(* IEC 61131-3 sources: sis-interlock-demo/pytests/golden/mini/tests/POUs/Generated/FB_CemGen01_Test, 24 files *)

(* ---- FB_CemGen01_Test.decl.st ---- *)
// AUTO-GENERATED by cemgen 1.0.0 — не редактировать: правьте матрицу и запустите
//   python -m cemgen generate <файл матрицы .csv или .xlsx>
// Матрица: TEST-U301-CEM, объект U-301, ревизия 1 от 2026-10-16, SHA-256 сетки 9067fda96ae55e67
// Назначение: набор coUnit: сценарии по матрице TEST-U301-CEM, тесты 1–24 (DESIGN.md, 12.4).
//             Ожидаемые значения — эталонная модель cemgen. Стенд FB_SisHarness — по экземпляру на
//             тест.
// Автор:      pytest; код — генератор cemgen
// Версия:     1.0.0
// Документ:   docs/DESIGN.md, раздел «10. Генератор cemgen»; docs/cause_effect_matrix.md
// ВНИМАНИЕ:   код демонстрационный и не предназначен для систем безопасности. Реальная ПАЗ требует
//             определения SIL, сертифицированных аппаратных и программных средств и валидации по
//             ГОСТ Р МЭК 61511.
FUNCTION_BLOCK FB_CemGen01_Test EXTENDS coUnit.FB_TestSuite
VAR
    fbH001 : FB_SisHarness;   // Matrix_TSH301Demand_TripsOwnEffects
    fbH002 : FB_SisHarness;   // Matrix_TSH301Delay_TripsExactlyAtDelay
    fbH003 : FB_SisHarness;   // Matrix_TSH301Override_Denied
    fbH004 : FB_SisHarness;   // Matrix_TSH301Reset_OnlyAfterClear
    fbH005 : FB_SisHarness;   // Matrix_TSH301ChannelInvalid_MatchesPolicy
    fbH006 : FB_SisHarness;   // Matrix_TSH301Bypass_Denied
    fbH007 : FB_SisHarness;   // Matrix_PSL302Demand_TripsOwnEffects
    fbH008 : FB_SisHarness;   // Matrix_PSL302Override_ExpiresThenTrips
    fbH009 : FB_SisHarness;   // Matrix_PSL302Override_ClearsAfterConfirm
    fbH010 : FB_SisHarness;   // Matrix_PSL302Override_DemandBackRestartsConfirm
    fbH011 : FB_SisHarness;   // Matrix_PSL302Override_ExpiryBoundsConfirm
    fbH012 : FB_SisHarness;   // Matrix_PSL302Reset_OnlyAfterClear
    fbH013 : FB_SisHarness;   // Matrix_PSL302ChannelInvalid_MatchesPolicy
    fbH014 : FB_SisHarness;   // Matrix_PSL302Bypass_ExpiresBackToVoting
    fbH015 : FB_SisHarness;   // Matrix_XS303Demand_TripsOwnEffects
    fbH016 : FB_SisHarness;   // Matrix_XS303Delay_TripsExactlyAtDelay
    fbH017 : FB_SisHarness;   // Matrix_XS303Override_Denied
    fbH018 : FB_SisHarness;   // Matrix_XS303Reset_OnlyAfterClear
    fbH019 : FB_SisHarness;   // Matrix_FirstOutTSH301ThenPSL302_RecordsFirst
    fbH020 : FB_SisHarness;   // Matrix_FirstOutPSL302ThenXS303_RecordsFirst
    fbH021 : FB_SisHarness;   // Matrix_FirstOutXS303ThenTSH301_RecordsFirst
    fbH022 : FB_SisHarness;   // Matrix_Start_EnergizedWithoutReset
    fbH023 : FB_SisHarness;   // Matrix_FirstOutSimultaneous_LowestIndex
    fbH024 : FB_SisHarness;   // Matrix_GeneratedCfg_PassesChecks
END_VAR

(* ---- FirstOutPSL302ThenXS303RecordsFirst.method.decl.st ---- *)
// AUTO-GENERATED by cemgen 1.0.0 — не редактировать: правьте матрицу и запустите
//   python -m cemgen generate <файл матрицы .csv или .xlsx>
// Матрица: TEST-U301-CEM, объект U-301, ревизия 1 от 2026-10-16, SHA-256 сетки 9067fda96ae55e67
// Назначение: тест Matrix_FirstOutPSL302ThenXS303_RecordsFirst набора FB_CemGen01_Test (сценарий по
//             матрице, DESIGN.md, 12.4).
// Автор:      pytest; код — генератор cemgen
// Версия:     1.0.0
// Документ:   docs/DESIGN.md, раздел «10. Генератор cemgen»; docs/cause_effect_matrix.md
// ВНИМАНИЕ:   код демонстрационный и не предназначен для систем безопасности. Реальная ПАЗ требует
//             определения SIL, сертифицированных аппаратных и программных средств и валидации по
//             ГОСТ Р МЭК 61511.
// Первопричина: требование PSL302, фиксация через 0 с; затем требование XS303, фиксация через 500 мс →
// первопричина PSL302, в маске первопричины только PSL302, ltFirstOut — момент фиксации PSL302, XS303
// — среди зафиксированных.
METHOD PRIVATE FirstOutPSL302ThenXS303RecordsFirst
VAR
    xArmed : BOOL;    // стенд взведён: все следствия под напряжением после сброса
    ltT0   : LTIME;   // момент t0 по подменному времени стенда
END_VAR

(* ---- FirstOutSimultaneousLowestIndex.method.decl.st ---- *)
// AUTO-GENERATED by cemgen 1.0.0 — не редактировать: правьте матрицу и запустите
//   python -m cemgen generate <файл матрицы .csv или .xlsx>
// Матрица: TEST-U301-CEM, объект U-301, ревизия 1 от 2026-10-16, SHA-256 сетки 9067fda96ae55e67
// Назначение: тест Matrix_FirstOutSimultaneous_LowestIndex набора FB_CemGen01_Test (сценарий по
//             матрице, DESIGN.md, 12.4).
// Автор:      pytest; код — генератор cemgen
// Версия:     1.0.0
// Документ:   docs/DESIGN.md, раздел «10. Генератор cemgen»; docs/cause_effect_matrix.md
// ВНИМАНИЕ:   код демонстрационный и не предназначен для систем безопасности. Реальная ПАЗ требует
//             определения SIL, сертифицированных аппаратных и программных средств и валидации по
//             ГОСТ Р МЭК 61511.
// Одновременная фиксация TSH301 и PSL302 (без общих каналов) в одном вызове: требования подаются со
// сдвигом на разницу задержек → первопричина — младшая причина, в маске первопричины обе.
METHOD PRIVATE FirstOutSimultaneousLowestIndex
VAR
    xArmed : BOOL;   // стенд взведён: все следствия под напряжением после сброса
END_VAR

(* ---- FirstOutTSH301ThenPSL302RecordsFirst.method.decl.st ---- *)
// AUTO-GENERATED by cemgen 1.0.0 — не редактировать: правьте матрицу и запустите
//   python -m cemgen generate <файл матрицы .csv или .xlsx>
// Матрица: TEST-U301-CEM, объект U-301, ревизия 1 от 2026-10-16, SHA-256 сетки 9067fda96ae55e67
// Назначение: тест Matrix_FirstOutTSH301ThenPSL302_RecordsFirst набора FB_CemGen01_Test (сценарий
//             по матрице, DESIGN.md, 12.4).
// Автор:      pytest; код — генератор cemgen
// Версия:     1.0.0
// Документ:   docs/DESIGN.md, раздел «10. Генератор cemgen»; docs/cause_effect_matrix.md
// ВНИМАНИЕ:   код демонстрационный и не предназначен для систем безопасности. Реальная ПАЗ требует
//             определения SIL, сертифицированных аппаратных и программных средств и валидации по
//             ГОСТ Р МЭК 61511.
// Первопричина: требование TSH301, фиксация через 1 с; затем требование PSL302, фиксация через 0 с →
// первопричина TSH301, в маске первопричины только TSH301, ltFirstOut — момент фиксации TSH301, PSL302
// — среди зафиксированных.
METHOD PRIVATE FirstOutTSH301ThenPSL302RecordsFirst
VAR
    xArmed : BOOL;    // стенд взведён: все следствия под напряжением после сброса
    ltT0   : LTIME;   // момент t0 по подменному времени стенда
END_VAR

(* ---- FirstOutXS303ThenTSH301RecordsFirst.method.decl.st ---- *)
// AUTO-GENERATED by cemgen 1.0.0 — не редактировать: правьте матрицу и запустите
//   python -m cemgen generate <файл матрицы .csv или .xlsx>
// Матрица: TEST-U301-CEM, объект U-301, ревизия 1 от 2026-10-16, SHA-256 сетки 9067fda96ae55e67
// Назначение: тест Matrix_FirstOutXS303ThenTSH301_RecordsFirst набора FB_CemGen01_Test (сценарий по
//             матрице, DESIGN.md, 12.4).
// Автор:      pytest; код — генератор cemgen
// Версия:     1.0.0
// Документ:   docs/DESIGN.md, раздел «10. Генератор cemgen»; docs/cause_effect_matrix.md
// ВНИМАНИЕ:   код демонстрационный и не предназначен для систем безопасности. Реальная ПАЗ требует
//             определения SIL, сертифицированных аппаратных и программных средств и валидации по
//             ГОСТ Р МЭК 61511.
// Первопричина: требование XS303, фиксация через 500 мс; затем требование TSH301, фиксация через 1 с →
// первопричина XS303, в маске первопричины только XS303, ltFirstOut — момент фиксации XS303, TSH301 —
// среди зафиксированных.
METHOD PRIVATE FirstOutXS303ThenTSH301RecordsFirst
VAR
    xArmed : BOOL;    // стенд взведён: все следствия под напряжением после сброса
    ltT0   : LTIME;   // момент t0 по подменному времени стенда
END_VAR

(* ---- GeneratedCfgPassesChecks.method.decl.st ---- *)
// AUTO-GENERATED by cemgen 1.0.0 — не редактировать: правьте матрицу и запустите
//   python -m cemgen generate <файл матрицы .csv или .xlsx>
// Матрица: TEST-U301-CEM, объект U-301, ревизия 1 от 2026-10-16, SHA-256 сетки 9067fda96ae55e67
// Назначение: тест Matrix_GeneratedCfg_PassesChecks набора FB_CemGen01_Test (сценарий по матрице,
//             DESIGN.md, 12.4).
// Автор:      pytest; код — генератор cemgen
// Версия:     1.0.0
// Документ:   docs/DESIGN.md, раздел «10. Генератор cemgen»; docs/cause_effect_matrix.md
// ВНИМАНИЕ:   код демонстрационный и не предназначен для систем безопасности. Реальная ПАЗ требует
//             определения SIL, сертифицированных аппаратных и программных средств и валидации по
//             ГОСТ Р МЭК 61511.
// Сгенерированная конфигурация: F_CemCrc(CEM_CFG) = 16#0F15 = CEM_CFG.wMatrixCrc, F_CemCheckCfg без
// ошибок; после взвода нет ошибок конфигурации у матрицы и у групп голосования.
METHOD PRIVATE GeneratedCfgPassesChecks
VAR
    stCfg  : ST_CemCfg;      // копия GVL_SisCfg.CEM_CFG
    wCrc   : WORD;           // CRC сгенерированной матрицы
    wErr   : WORD;           // биты ошибок конфигурации матрицы
    xArmed : BOOL;           // стенд взведён: все следствия под напряжением после сброса
    stVs   : ST_VotingSts;   // копия состояния группы голосования
END_VAR

(* ---- PSL302BypassExpiresBackToVoting.method.decl.st ---- *)
// AUTO-GENERATED by cemgen 1.0.0 — не редактировать: правьте матрицу и запустите
//   python -m cemgen generate <файл матрицы .csv или .xlsx>
// Матрица: TEST-U301-CEM, объект U-301, ревизия 1 от 2026-10-16, SHA-256 сетки 9067fda96ae55e67
// Назначение: тест Matrix_PSL302Bypass_ExpiresBackToVoting набора FB_CemGen01_Test (сценарий по
//             матрице, DESIGN.md, 12.4).
// Автор:      pytest; код — генератор cemgen
// Версия:     1.0.0
// Документ:   docs/DESIGN.md, раздел «10. Генератор cemgen»; docs/cause_effect_matrix.md
// ВНИМАНИЕ:   код демонстрационный и не предназначен для систем безопасности. Реальная ПАЗ требует
//             определения SIL, сертифицированных аппаратных и программных средств и валидации по
//             ГОСТ Р МЭК 61511.
// Причина 2 PSL302: ключ разрешения байпасов, байпас PS302A → Active; канал недостоверен → Bypassed,
// не сработало; на t0 + 1 ч − шаг — Active; ровно на t0 + 1 ч — Expired, BypassExpired, канал Invalid;
// далее — по эталонной модели.
METHOD PRIVATE PSL302BypassExpiresBackToVoting
VAR
    xArmed : BOOL;           // стенд взведён: все следствия под напряжением после сброса
    stVs   : ST_VotingSts;   // копия состояния группы голосования
END_VAR

(* ---- PSL302ChannelInvalidMatchesPolicy.method.decl.st ---- *)
// AUTO-GENERATED by cemgen 1.0.0 — не редактировать: правьте матрицу и запустите
//   python -m cemgen generate <файл матрицы .csv или .xlsx>
// Матрица: TEST-U301-CEM, объект U-301, ревизия 1 от 2026-10-16, SHA-256 сетки 9067fda96ae55e67
// Назначение: тест Matrix_PSL302ChannelInvalid_MatchesPolicy набора FB_CemGen01_Test (сценарий по
//             матрице, DESIGN.md, 12.4).
// Автор:      pytest; код — генератор cemgen
// Версия:     1.0.0
// Документ:   docs/DESIGN.md, раздел «10. Генератор cemgen»; docs/cause_effect_matrix.md
// ВНИМАНИЕ:   код демонстрационный и не предназначен для систем безопасности. Реальная ПАЗ требует
//             определения SIL, сертифицированных аппаратных и программных средств и валидации по
//             ГОСТ Р МЭК 61511.
// Причина 2 PSL302 (2oo2, VoteTrip): канал PS302A недостоверен → действующая схема и срабатывание по
// политике деградации; если не сработало — требование на PS302B → по эталонной модели.
METHOD PRIVATE PSL302ChannelInvalidMatchesPolicy
VAR
    xArmed : BOOL;           // стенд взведён: все следствия под напряжением после сброса
    stVs   : ST_VotingSts;   // копия состояния группы голосования
END_VAR

(* ---- PSL302DemandTripsOwnEffects.method.decl.st ---- *)
// AUTO-GENERATED by cemgen 1.0.0 — не редактировать: правьте матрицу и запустите
//   python -m cemgen generate <файл матрицы .csv или .xlsx>
// Матрица: TEST-U301-CEM, объект U-301, ревизия 1 от 2026-10-16, SHA-256 сетки 9067fda96ae55e67
// Назначение: тест Matrix_PSL302Demand_TripsOwnEffects набора FB_CemGen01_Test (сценарий по
//             матрице, DESIGN.md, 12.4).
// Автор:      pytest; код — генератор cemgen
// Версия:     1.0.0
// Документ:   docs/DESIGN.md, раздел «10. Генератор cemgen»; docs/cause_effect_matrix.md
// ВНИМАНИЕ:   код демонстрационный и не предназначен для систем безопасности. Реальная ПАЗ требует
//             определения SIL, сертифицированных аппаратных и программных средств и валидации по
//             ГОСТ Р МЭК 61511.
// Причина 2 PSL302 (2oo2, задержка 0 с): требование PS302A, PS302B = 0 отключает XV301, M302;
// остальные следствия под напряжением; первопричина PSL302.
METHOD PRIVATE PSL302DemandTripsOwnEffects
VAR
    xArmed : BOOL;   // стенд взведён: все следствия под напряжением после сброса
END_VAR

(* ---- PSL302OverrideClearsAfterConfirm.method.decl.st ---- *)
// AUTO-GENERATED by cemgen 1.0.0 — не редактировать: правьте матрицу и запустите
//   python -m cemgen generate <файл матрицы .csv или .xlsx>
// Матрица: TEST-U301-CEM, объект U-301, ревизия 1 от 2026-10-16, SHA-256 сетки 9067fda96ae55e67
// Назначение: тест Matrix_PSL302Override_ClearsAfterConfirm набора FB_CemGen01_Test (сценарий по
//             матрице, DESIGN.md, 12.4).
// Автор:      pytest; код — генератор cemgen
// Версия:     1.0.0
// Документ:   docs/DESIGN.md, раздел «10. Генератор cemgen»; docs/cause_effect_matrix.md
// ВНИМАНИЕ:   код демонстрационный и не предназначен для систем безопасности. Реальная ПАЗ требует
//             определения SIL, сертифицированных аппаратных и программных средств и валидации по
//             ГОСТ Р МЭК 61511.
// Причина 2 PSL302: пусковой обход и требование в t0; норма с t1 = t0 + шаг; на t1 + 30 с − шаг обход
// действует; ровно на t1 + 30 с (подтверждение нормы) — OverrideCleared, обхода нет, причина не
// зафиксирована, следствия под напряжением (R-12).
METHOD PRIVATE PSL302OverrideClearsAfterConfirm
VAR
    xArmed : BOOL;   // стенд взведён: все следствия под напряжением после сброса
END_VAR

(* ---- PSL302OverrideDemandBackRestartsConfirm.method.decl.st ---- *)
// AUTO-GENERATED by cemgen 1.0.0 — не редактировать: правьте матрицу и запустите
//   python -m cemgen generate <файл матрицы .csv или .xlsx>
// Матрица: TEST-U301-CEM, объект U-301, ревизия 1 от 2026-10-16, SHA-256 сетки 9067fda96ae55e67
// Назначение: тест Matrix_PSL302Override_DemandBackRestartsConfirm набора FB_CemGen01_Test
//             (сценарий по матрице, DESIGN.md, 12.4).
// Автор:      pytest; код — генератор cemgen
// Версия:     1.0.0
// Документ:   docs/DESIGN.md, раздел «10. Генератор cemgen»; docs/cause_effect_matrix.md
// ВНИМАНИЕ:   код демонстрационный и не предназначен для систем безопасности. Реальная ПАЗ требует
//             определения SIL, сертифицированных аппаратных и программных средств и валидации по
//             ГОСТ Р МЭК 61511.
// Причина 2 PSL302: пусковой обход и требование в t0; норма с t1; ровно на t1 + 30 с, когда обход
// снялся бы, требование снова — обход действует, подтверждение нормы сброшено; норма с t2; на t2 + 30
// с − шаг обход действует; на t2 + 30 с — OverrideCleared.
METHOD PRIVATE PSL302OverrideDemandBackRestartsConfirm
VAR
    xArmed : BOOL;   // стенд взведён: все следствия под напряжением после сброса
END_VAR

(* ---- PSL302OverrideExpiresThenTrips.method.decl.st ---- *)
// AUTO-GENERATED by cemgen 1.0.0 — не редактировать: правьте матрицу и запустите
//   python -m cemgen generate <файл матрицы .csv или .xlsx>
// Матрица: TEST-U301-CEM, объект U-301, ревизия 1 от 2026-10-16, SHA-256 сетки 9067fda96ae55e67
// Назначение: тест Matrix_PSL302Override_ExpiresThenTrips набора FB_CemGen01_Test (сценарий по
//             матрице, DESIGN.md, 12.4).
// Автор:      pytest; код — генератор cemgen
// Версия:     1.0.0
// Документ:   docs/DESIGN.md, раздел «10. Генератор cemgen»; docs/cause_effect_matrix.md
// ВНИМАНИЕ:   код демонстрационный и не предназначен для систем безопасности. Реальная ПАЗ требует
//             определения SIL, сертифицированных аппаратных и программных средств и валидации по
//             ГОСТ Р МЭК 61511.
// Причина 2 PSL302: ключ разрешения обходов, запрос пускового обхода и требование в одном вызове t0;
// до t0 + 10 мин − шаг обход действует, причина не зафиксирована; ровно на t0 + 10 мин —
// OverrideExpired, фиксация, первопричина PSL302.
METHOD PRIVATE PSL302OverrideExpiresThenTrips
VAR
    xArmed : BOOL;   // стенд взведён: все следствия под напряжением после сброса
END_VAR

(* ---- PSL302OverrideExpiryBoundsConfirm.method.decl.st ---- *)
// AUTO-GENERATED by cemgen 1.0.0 — не редактировать: правьте матрицу и запустите
//   python -m cemgen generate <файл матрицы .csv или .xlsx>
// Матрица: TEST-U301-CEM, объект U-301, ревизия 1 от 2026-10-16, SHA-256 сетки 9067fda96ae55e67
// Назначение: тест Matrix_PSL302Override_ExpiryBoundsConfirm набора FB_CemGen01_Test (сценарий по
//             матрице, DESIGN.md, 12.4).
// Автор:      pytest; код — генератор cemgen
// Версия:     1.0.0
// Документ:   docs/DESIGN.md, раздел «10. Генератор cemgen»; docs/cause_effect_matrix.md
// ВНИМАНИЕ:   код демонстрационный и не предназначен для систем безопасности. Реальная ПАЗ требует
//             определения SIL, сертифицированных аппаратных и программных средств и валидации по
//             ГОСТ Р МЭК 61511.
// Причина 2 PSL302: пусковой обход и требование в t0; норма с t0 + 9 мин 30 с + шаг — подтверждение
// (30 с) закончилось бы после срока; на t0 + 10 мин − шаг обход действует; ровно на t0 + 10 мин —
// OverrideExpired (срок — верхняя граница), OverrideCleared нет, причина не зафиксирована (требования
// нет).
METHOD PRIVATE PSL302OverrideExpiryBoundsConfirm
VAR
    xArmed : BOOL;   // стенд взведён: все следствия под напряжением после сброса
END_VAR

(* ---- PSL302ResetOnlyAfterClear.method.decl.st ---- *)
// AUTO-GENERATED by cemgen 1.0.0 — не редактировать: правьте матрицу и запустите
//   python -m cemgen generate <файл матрицы .csv или .xlsx>
// Матрица: TEST-U301-CEM, объект U-301, ревизия 1 от 2026-10-16, SHA-256 сетки 9067fda96ae55e67
// Назначение: тест Matrix_PSL302Reset_OnlyAfterClear набора FB_CemGen01_Test (сценарий по матрице,
//             DESIGN.md, 12.4).
// Автор:      pytest; код — генератор cemgen
// Версия:     1.0.0
// Документ:   docs/DESIGN.md, раздел «10. Генератор cemgen»; docs/cause_effect_matrix.md
// ВНИМАНИЕ:   код демонстрационный и не предназначен для систем безопасности. Реальная ПАЗ требует
//             определения SIL, сертифицированных аппаратных и программных средств и валидации по
//             ГОСТ Р МЭК 61511.
// Причина 2 PSL302: срабатывание; сброс при требовании → ResetDenied, блокирует PSL302, следствия
// обесточены; норма → следствия всё ещё обесточены (фиксация); сброс → все следствия под напряжением.
METHOD PRIVATE PSL302ResetOnlyAfterClear
VAR
    xArmed : BOOL;          // стенд взведён: все следствия под напряжением после сброса
    stEv   : ST_SisEvent;   // последнее событие журнала
END_VAR

(* ---- TSH301BypassDenied.method.decl.st ---- *)
// AUTO-GENERATED by cemgen 1.0.0 — не редактировать: правьте матрицу и запустите
//   python -m cemgen generate <файл матрицы .csv или .xlsx>
// Матрица: TEST-U301-CEM, объект U-301, ревизия 1 от 2026-10-16, SHA-256 сетки 9067fda96ae55e67
// Назначение: тест Matrix_TSH301Bypass_Denied набора FB_CemGen01_Test (сценарий по матрице,
//             DESIGN.md, 12.4).
// Автор:      pytest; код — генератор cemgen
// Версия:     1.0.0
// Документ:   docs/DESIGN.md, раздел «10. Генератор cemgen»; docs/cause_effect_matrix.md
// ВНИМАНИЕ:   код демонстрационный и не предназначен для систем безопасности. Реальная ПАЗ требует
//             определения SIL, сертифицированных аппаратных и программных средств и валидации по
//             ГОСТ Р МЭК 61511.
// Причина 1 TSH301: байпас запрещён (bypass_max = 0); ключ разрешения байпасов, запрос байпаса TT301 →
// Denied, событие BypassDenied с номером канала.
METHOD PRIVATE TSH301BypassDenied
VAR
    xArmed : BOOL;           // стенд взведён: все следствия под напряжением после сброса
    stVs   : ST_VotingSts;   // копия состояния группы голосования
    stEv   : ST_SisEvent;    // последнее событие журнала
END_VAR

(* ---- TSH301ChannelInvalidMatchesPolicy.method.decl.st ---- *)
// AUTO-GENERATED by cemgen 1.0.0 — не редактировать: правьте матрицу и запустите
//   python -m cemgen generate <файл матрицы .csv или .xlsx>
// Матрица: TEST-U301-CEM, объект U-301, ревизия 1 от 2026-10-16, SHA-256 сетки 9067fda96ae55e67
// Назначение: тест Matrix_TSH301ChannelInvalid_MatchesPolicy набора FB_CemGen01_Test (сценарий по
//             матрице, DESIGN.md, 12.4).
// Автор:      pytest; код — генератор cemgen
// Версия:     1.0.0
// Документ:   docs/DESIGN.md, раздел «10. Генератор cemgen»; docs/cause_effect_matrix.md
// ВНИМАНИЕ:   код демонстрационный и не предназначен для систем безопасности. Реальная ПАЗ требует
//             определения SIL, сертифицированных аппаратных и программных средств и валидации по
//             ГОСТ Р МЭК 61511.
// Причина 1 TSH301 (1oo1, VoteTrip): канал TT301 недостоверен → действующая схема и срабатывание по
// политике деградации; если не сработало — требование на втором канале → по эталонной модели.
METHOD PRIVATE TSH301ChannelInvalidMatchesPolicy
VAR
    xArmed : BOOL;           // стенд взведён: все следствия под напряжением после сброса
    stVs   : ST_VotingSts;   // копия состояния группы голосования
END_VAR

(* ---- TSH301DelayTripsExactlyAtDelay.method.decl.st ---- *)
// AUTO-GENERATED by cemgen 1.0.0 — не редактировать: правьте матрицу и запустите
//   python -m cemgen generate <файл матрицы .csv или .xlsx>
// Матрица: TEST-U301-CEM, объект U-301, ревизия 1 от 2026-10-16, SHA-256 сетки 9067fda96ae55e67
// Назначение: тест Matrix_TSH301Delay_TripsExactlyAtDelay набора FB_CemGen01_Test (сценарий по
//             матрице, DESIGN.md, 12.4).
// Автор:      pytest; код — генератор cemgen
// Версия:     1.0.0
// Документ:   docs/DESIGN.md, раздел «10. Генератор cemgen»; docs/cause_effect_matrix.md
// ВНИМАНИЕ:   код демонстрационный и не предназначен для систем безопасности. Реальная ПАЗ требует
//             определения SIL, сертифицированных аппаратных и программных средств и валидации по
//             ГОСТ Р МЭК 61511.
// Причина 1 TSH301: требование в t0; на t0 + 1 с − шаг не зафиксирована, следствия под напряжением;
// ровно на t0 + 1 с — зафиксирована, ltFirstOut = t0 + задержка.
METHOD PRIVATE TSH301DelayTripsExactlyAtDelay
VAR
    xArmed : BOOL;    // стенд взведён: все следствия под напряжением после сброса
    ltT0   : LTIME;   // момент t0 по подменному времени стенда
END_VAR

(* ---- TSH301DemandTripsOwnEffects.method.decl.st ---- *)
// AUTO-GENERATED by cemgen 1.0.0 — не редактировать: правьте матрицу и запустите
//   python -m cemgen generate <файл матрицы .csv или .xlsx>
// Матрица: TEST-U301-CEM, объект U-301, ревизия 1 от 2026-10-16, SHA-256 сетки 9067fda96ae55e67
// Назначение: тест Matrix_TSH301Demand_TripsOwnEffects набора FB_CemGen01_Test (сценарий по
//             матрице, DESIGN.md, 12.4).
// Автор:      pytest; код — генератор cemgen
// Версия:     1.0.0
// Документ:   docs/DESIGN.md, раздел «10. Генератор cemgen»; docs/cause_effect_matrix.md
// ВНИМАНИЕ:   код демонстрационный и не предназначен для систем безопасности. Реальная ПАЗ требует
//             определения SIL, сертифицированных аппаратных и программных средств и валидации по
//             ГОСТ Р МЭК 61511.
// Причина 1 TSH301 (1oo1, задержка 1 с): требование TT301 = 16,96 мА (81 °C; уставка ≥ 80 °C)
// отключает XV301; остальные следствия под напряжением; первопричина TSH301.
METHOD PRIVATE TSH301DemandTripsOwnEffects
VAR
    xArmed : BOOL;   // стенд взведён: все следствия под напряжением после сброса
END_VAR

(* ---- TSH301OverrideDenied.method.decl.st ---- *)
// AUTO-GENERATED by cemgen 1.0.0 — не редактировать: правьте матрицу и запустите
//   python -m cemgen generate <файл матрицы .csv или .xlsx>
// Матрица: TEST-U301-CEM, объект U-301, ревизия 1 от 2026-10-16, SHA-256 сетки 9067fda96ae55e67
// Назначение: тест Matrix_TSH301Override_Denied набора FB_CemGen01_Test (сценарий по матрице,
//             DESIGN.md, 12.4).
// Автор:      pytest; код — генератор cemgen
// Версия:     1.0.0
// Документ:   docs/DESIGN.md, раздел «10. Генератор cemgen»; docs/cause_effect_matrix.md
// ВНИМАНИЕ:   код демонстрационный и не предназначен для систем безопасности. Реальная ПАЗ требует
//             определения SIL, сертифицированных аппаратных и программных средств и валидации по
//             ГОСТ Р МЭК 61511.
// Причина 1 TSH301 без разрешённого обхода: ключ разрешения обходов, запрос → последнее событие
// OverrideDenied, обхода нет; требование → срабатывание после задержки.
METHOD PRIVATE TSH301OverrideDenied
VAR
    xArmed : BOOL;          // стенд взведён: все следствия под напряжением после сброса
    stEv   : ST_SisEvent;   // последнее событие журнала
END_VAR

(* ---- TSH301ResetOnlyAfterClear.method.decl.st ---- *)
// AUTO-GENERATED by cemgen 1.0.0 — не редактировать: правьте матрицу и запустите
//   python -m cemgen generate <файл матрицы .csv или .xlsx>
// Матрица: TEST-U301-CEM, объект U-301, ревизия 1 от 2026-10-16, SHA-256 сетки 9067fda96ae55e67
// Назначение: тест Matrix_TSH301Reset_OnlyAfterClear набора FB_CemGen01_Test (сценарий по матрице,
//             DESIGN.md, 12.4).
// Автор:      pytest; код — генератор cemgen
// Версия:     1.0.0
// Документ:   docs/DESIGN.md, раздел «10. Генератор cemgen»; docs/cause_effect_matrix.md
// ВНИМАНИЕ:   код демонстрационный и не предназначен для систем безопасности. Реальная ПАЗ требует
//             определения SIL, сертифицированных аппаратных и программных средств и валидации по
//             ГОСТ Р МЭК 61511.
// Причина 1 TSH301: срабатывание; сброс при требовании → ResetDenied, блокирует TSH301, следствия
// обесточены; норма → следствия всё ещё обесточены (фиксация); сброс → все следствия под напряжением.
METHOD PRIVATE TSH301ResetOnlyAfterClear
VAR
    xArmed : BOOL;          // стенд взведён: все следствия под напряжением после сброса
    stEv   : ST_SisEvent;   // последнее событие журнала
END_VAR

(* ---- XS303DelayTripsExactlyAtDelay.method.decl.st ---- *)
// AUTO-GENERATED by cemgen 1.0.0 — не редактировать: правьте матрицу и запустите
//   python -m cemgen generate <файл матрицы .csv или .xlsx>
// Матрица: TEST-U301-CEM, объект U-301, ревизия 1 от 2026-10-16, SHA-256 сетки 9067fda96ae55e67
// Назначение: тест Matrix_XS303Delay_TripsExactlyAtDelay набора FB_CemGen01_Test (сценарий по
//             матрице, DESIGN.md, 12.4).
// Автор:      pytest; код — генератор cemgen
// Версия:     1.0.0
// Документ:   docs/DESIGN.md, раздел «10. Генератор cemgen»; docs/cause_effect_matrix.md
// ВНИМАНИЕ:   код демонстрационный и не предназначен для систем безопасности. Реальная ПАЗ требует
//             определения SIL, сертифицированных аппаратных и программных средств и валидации по
//             ГОСТ Р МЭК 61511.
// Причина 3 XS303: требование в t0; на t0 + 500 мс − шаг не зафиксирована, следствия под напряжением;
// ровно на t0 + 500 мс — зафиксирована, ltFirstOut = t0 + задержка.
METHOD PRIVATE XS303DelayTripsExactlyAtDelay
VAR
    xArmed : BOOL;    // стенд взведён: все следствия под напряжением после сброса
    ltT0   : LTIME;   // момент t0 по подменному времени стенда
END_VAR

(* ---- XS303DemandTripsOwnEffects.method.decl.st ---- *)
// AUTO-GENERATED by cemgen 1.0.0 — не редактировать: правьте матрицу и запустите
//   python -m cemgen generate <файл матрицы .csv или .xlsx>
// Матрица: TEST-U301-CEM, объект U-301, ревизия 1 от 2026-10-16, SHA-256 сетки 9067fda96ae55e67
// Назначение: тест Matrix_XS303Demand_TripsOwnEffects набора FB_CemGen01_Test (сценарий по матрице,
//             DESIGN.md, 12.4).
// Автор:      pytest; код — генератор cemgen
// Версия:     1.0.0
// Документ:   docs/DESIGN.md, раздел «10. Генератор cemgen»; docs/cause_effect_matrix.md
// ВНИМАНИЕ:   код демонстрационный и не предназначен для систем безопасности. Реальная ПАЗ требует
//             определения SIL, сертифицированных аппаратных и программных средств и валидации по
//             ГОСТ Р МЭК 61511.
// Причина 3 XS303 (—, задержка 500 мс): требование XS303 = 1 отключает M302; остальные следствия под
// напряжением; первопричина XS303.
METHOD PRIVATE XS303DemandTripsOwnEffects
VAR
    xArmed : BOOL;   // стенд взведён: все следствия под напряжением после сброса
END_VAR

(* ---- XS303OverrideDenied.method.decl.st ---- *)
// AUTO-GENERATED by cemgen 1.0.0 — не редактировать: правьте матрицу и запустите
//   python -m cemgen generate <файл матрицы .csv или .xlsx>
// Матрица: TEST-U301-CEM, объект U-301, ревизия 1 от 2026-10-16, SHA-256 сетки 9067fda96ae55e67
// Назначение: тест Matrix_XS303Override_Denied набора FB_CemGen01_Test (сценарий по матрице,
//             DESIGN.md, 12.4).
// Автор:      pytest; код — генератор cemgen
// Версия:     1.0.0
// Документ:   docs/DESIGN.md, раздел «10. Генератор cemgen»; docs/cause_effect_matrix.md
// ВНИМАНИЕ:   код демонстрационный и не предназначен для систем безопасности. Реальная ПАЗ требует
//             определения SIL, сертифицированных аппаратных и программных средств и валидации по
//             ГОСТ Р МЭК 61511.
// Причина 3 XS303 без разрешённого обхода: ключ разрешения обходов, запрос → последнее событие
// OverrideDenied, обхода нет; требование → срабатывание после задержки.
METHOD PRIVATE XS303OverrideDenied
VAR
    xArmed : BOOL;          // стенд взведён: все следствия под напряжением после сброса
    stEv   : ST_SisEvent;   // последнее событие журнала
END_VAR

(* ---- XS303ResetOnlyAfterClear.method.decl.st ---- *)
// AUTO-GENERATED by cemgen 1.0.0 — не редактировать: правьте матрицу и запустите
//   python -m cemgen generate <файл матрицы .csv или .xlsx>
// Матрица: TEST-U301-CEM, объект U-301, ревизия 1 от 2026-10-16, SHA-256 сетки 9067fda96ae55e67
// Назначение: тест Matrix_XS303Reset_OnlyAfterClear набора FB_CemGen01_Test (сценарий по матрице,
//             DESIGN.md, 12.4).
// Автор:      pytest; код — генератор cemgen
// Версия:     1.0.0
// Документ:   docs/DESIGN.md, раздел «10. Генератор cemgen»; docs/cause_effect_matrix.md
// ВНИМАНИЕ:   код демонстрационный и не предназначен для систем безопасности. Реальная ПАЗ требует
//             определения SIL, сертифицированных аппаратных и программных средств и валидации по
//             ГОСТ Р МЭК 61511.
// Причина 3 XS303: срабатывание; сброс при требовании → ResetDenied, блокирует XS303, следствия
// обесточены; норма → следствия всё ещё обесточены (фиксация); сброс → все следствия под напряжением.
METHOD PRIVATE XS303ResetOnlyAfterClear
VAR
    xArmed : BOOL;          // стенд взведён: все следствия под напряжением после сброса
    stEv   : ST_SisEvent;   // последнее событие журнала
END_VAR
